// TIA Portal project "2026_09_21_Ciclo_L" (V15)

(* hardware
DEVICE "S7-1200 station_1"  S7-1200 Station
   slot 0: "Telaio di montaggio_0"  S7-1200 Rack  Rack  V1.0
   slot 1: "PLC_1"  CPU 1215C DC/DC/DC  6ES7 215-1AG40-0XB0  V4.2
*)

// ===== PLC "PLC_1"  CPU 1215C DC/DC/DC =====

VAR_GLOBAL   // PLC tag table "Tabella delle variabili standard"
   "IC" AT %I0.0 : Bool;   // Pulsante di inizio ciclo
   "FC" AT %I0.1 : Bool;   // Pulsante di fine ciclo
   "a0" AT %I0.2 : Bool;   // Fine corsa cilindro A chiuso
   "a1" AT %I0.3 : Bool;   // Fine corsa cilindro A aperto
   "b0" AT %I0.4 : Bool;   // Fine corsa cilindro B chiuso
   "b1" AT %I0.5 : Bool;   // Fine corsa cilindro B aperto
   "A+" AT %Q0.0 : Bool;   // Fase positiva cilindro A
   "A-" AT %Q0.1 : Bool;   // Fase negativa cilindro A
   "B+" AT %Q0.2 : Bool;   // Fase positiva cilindro B
   "B-" AT %Q0.3 : Bool;   // Fase negativa cilindro B
   "HL0" AT %Q0.4 : Bool;   // Lampada di segnalazione impianto spento
   "HL1" AT %Q0.5 : Bool;   // Lampada di segnalazione impianto acceso
   "P0" AT %M10.0 : Bool;   // Fase 0
   "P1" AT %M10.1 : Bool;   // Fase 1
   "P2" AT %M10.2 : Bool;   // Fase 2
   "P3" AT %M10.3 : Bool;   // Fase 3
   "P4" AT %M10.4 : Bool;   // Fase 4
   "IC_V" AT %M20.0 : Bool;   // Start virtuale
   "FC_V" AT %M20.1 : Bool;
   "a0_V" AT %M20.2 : Bool;
   "a1_V" AT %M20.3 : Bool;
   "b0_V" AT %M20.4 : Bool;
   "b1_V" AT %M20.5 : Bool;
END_VAR

FUNCTION "Controllo" : Void   // FC1, LAD
{ S7_Optimized_Access := 'TRUE' }
VERSION : 0.1
   VAR_TEMP   // added for the SCL form of the ladder/FBD networks
      _w1 : Bool;
   END_VAR
BEGIN

REGION Network 1: Fase 0
   // Alla pressione del pulsante di Start, si avvia il ciclo di lavoro (stato 1)
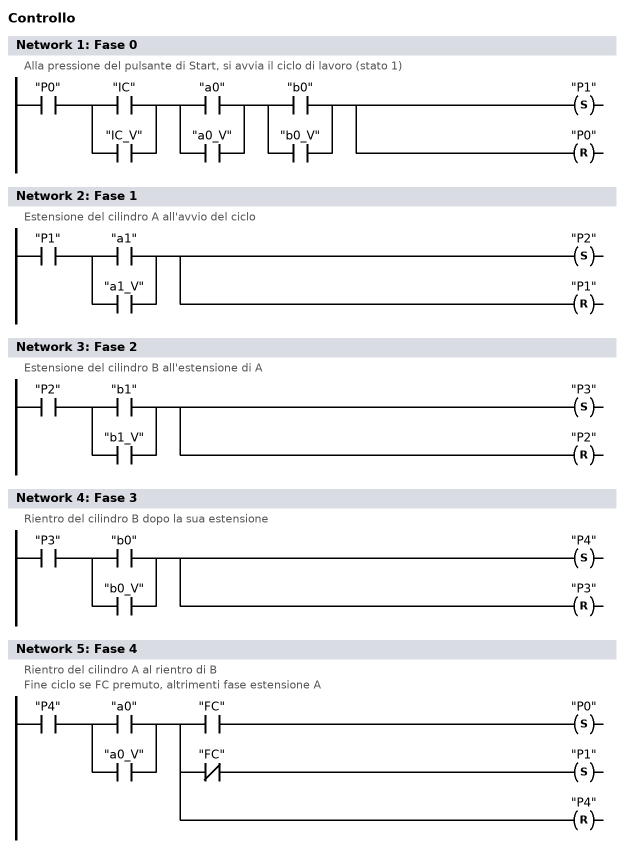
   RUNG wire#powerrail
      Contact( "P0" )
      wire#w1
      Contact( "IC" )
      wire#w2
      Contact( "a0" )
      wire#w3
      Contact( "b0" )
      wire#w4
      S_Coil( "P1" )
   END_RUNG
   RUNG wire#w1
      Contact( "IC_V" )
   END_RUNG wire#w2
   RUNG wire#w2
      Contact( "a0_V" )
   END_RUNG wire#w3
   RUNG wire#w3
      Contact( "b0_V" )
   END_RUNG wire#w4
   RUNG wire#w4
      R_Coil( "P0" )
   END_RUNG
   // the same network as SCL:
   IF "P0" AND ("IC" OR "IC_V") AND ("a0" OR "a0_V") AND ("b0" OR "b0_V") THEN
       "P1" := TRUE;
       "P0" := FALSE;
   END_IF;
END_REGION

REGION Network 2: Fase 1
   // Estensione del cilindro A all'avvio del ciclo
   RUNG wire#powerrail
      Contact( "P1" )
      wire#w1
      Contact( "a1" )
      wire#w2
      S_Coil( "P2" )
   END_RUNG
   RUNG wire#w1
      Contact( "a1_V" )
   END_RUNG wire#w2
   RUNG wire#w2
      R_Coil( "P1" )
   END_RUNG
   // the same network as SCL:
   IF "P1" AND ("a1" OR "a1_V") THEN
       "P2" := TRUE;
       "P1" := FALSE;
   END_IF;
END_REGION

REGION Network 3: Fase 2
   // Estensione del cilindro B all'estensione di A
   RUNG wire#powerrail
      Contact( "P2" )
      wire#w1
      Contact( "b1" )
      wire#w2
      S_Coil( "P3" )
   END_RUNG
   RUNG wire#w1
      Contact( "b1_V" )
   END_RUNG wire#w2
   RUNG wire#w2
      R_Coil( "P2" )
   END_RUNG
   // the same network as SCL:
   IF "P2" AND ("b1" OR "b1_V") THEN
       "P3" := TRUE;
       "P2" := FALSE;
   END_IF;
END_REGION

REGION Network 4: Fase 3
   // Rientro del cilindro B dopo la sua estensione
   RUNG wire#powerrail
      Contact( "P3" )
      wire#w1
      Contact( "b0" )
      wire#w2
      S_Coil( "P4" )
   END_RUNG
   RUNG wire#w1
      Contact( "b0_V" )
   END_RUNG wire#w2
   RUNG wire#w2
      R_Coil( "P3" )
   END_RUNG
   // the same network as SCL:
   IF "P3" AND ("b0" OR "b0_V") THEN
       "P4" := TRUE;
       "P3" := FALSE;
   END_IF;
END_REGION

REGION Network 5: Fase 4
   // Rientro del cilindro A al rientro di B
   // Fine ciclo se FC premuto, altrimenti fase estensione A
   RUNG wire#powerrail
      Contact( "P4" )
      wire#w1
      Contact( "a0" )
      wire#w2
      Contact( "FC" )
      S_Coil( "P0" )
   END_RUNG
   RUNG wire#w1
      Contact( "a0_V" )
   END_RUNG wire#w2
   RUNG wire#w2
      I_Contact( "FC" )
      S_Coil( "P1" )
   END_RUNG
   RUNG wire#w2
      R_Coil( "P4" )
   END_RUNG
   // the same network as SCL:
   #_w1 := "P4" AND ("a0" OR "a0_V");
   IF #_w1 AND "FC" THEN "P0" := TRUE; END_IF;
   IF #_w1 AND NOT "FC" THEN "P1" := TRUE; END_IF;
   IF #_w1 THEN "P4" := FALSE; END_IF;
END_REGION
END_FUNCTION

FUNCTION "Comando" : Void   // FC2, LAD
{ S7_Optimized_Access := 'TRUE' }
VERSION : 0.1
BEGIN

REGION Network 1: Lampada di segnalazione impianto spento
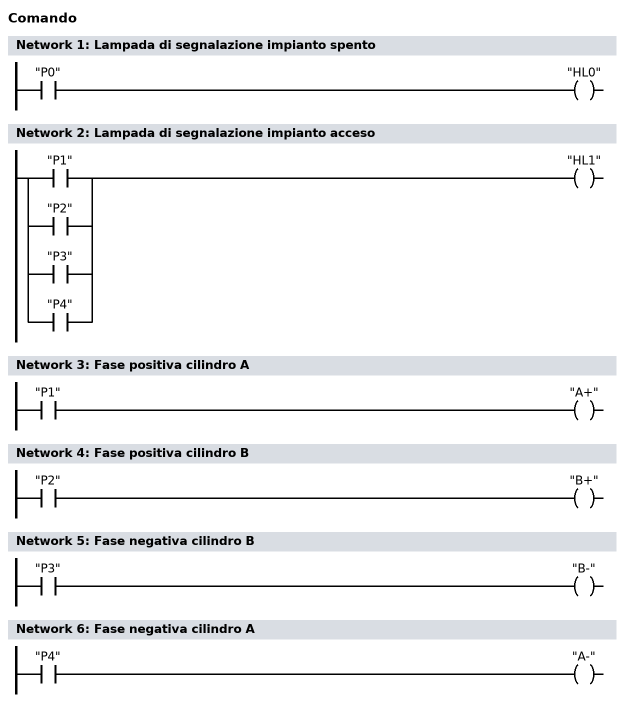
   RUNG wire#powerrail
      Contact( "P0" )
      Coil( "HL0" )
   END_RUNG
   // the same network as SCL:
   "HL0" := "P0";
END_REGION

REGION Network 2: Lampada di segnalazione impianto acceso
   RUNG wire#powerrail
      Contact( "P1" )
      wire#w1
      Coil( "HL1" )
   END_RUNG
   RUNG wire#powerrail
      Contact( "P2" )
   END_RUNG wire#w1
   RUNG wire#powerrail
      Contact( "P3" )
   END_RUNG wire#w1
   RUNG wire#powerrail
      Contact( "P4" )
   END_RUNG wire#w1
   // the same network as SCL:
   "HL1" := "P1" OR "P2" OR "P3" OR "P4";
END_REGION

REGION Network 3: Fase positiva cilindro A
   RUNG wire#powerrail
      Contact( "P1" )
      Coil( "A+" )
   END_RUNG
   // the same network as SCL:
   "A+" := "P1";
END_REGION

REGION Network 4: Fase positiva cilindro B
   RUNG wire#powerrail
      Contact( "P2" )
      Coil( "B+" )
   END_RUNG
   // the same network as SCL:
   "B+" := "P2";
END_REGION

REGION Network 5: Fase negativa cilindro B
   RUNG wire#powerrail
      Contact( "P3" )
      Coil( "B-" )
   END_RUNG
   // the same network as SCL:
   "B-" := "P3";
END_REGION

REGION Network 6: Fase negativa cilindro A
   RUNG wire#powerrail
      Contact( "P4" )
      Coil( "A-" )
   END_RUNG
   // the same network as SCL:
   "A-" := "P4";
END_REGION
END_FUNCTION

ORGANIZATION_BLOCK "Main"   // OB1, LAD, ProgramCycle
TITLE = "Main Program Sweep (Cycle)"
{ S7_Optimized_Access := 'TRUE' }
VERSION : 0.1
   VAR_INPUT
      Initial_Call : Bool;   // Initial call of this OB
      Remanence : Bool;   // =True, if remanent data are available
   END_VAR
BEGIN

REGION Network 1: FC Controllo
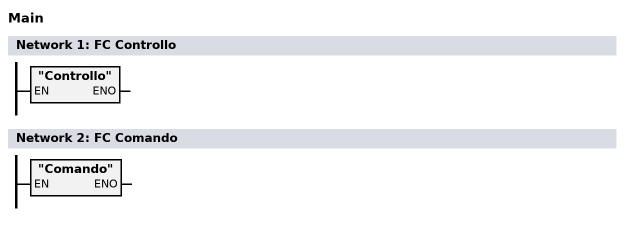
   RUNG wire#powerrail
      "Controllo"()
   END_RUNG
   // the same network as SCL:
   "Controllo"();
END_REGION

REGION Network 2: FC Comando
   RUNG wire#powerrail
      "Comando"()
   END_RUNG
   // the same network as SCL:
   "Comando"();
END_REGION
END_ORGANIZATION_BLOCK

ORGANIZATION_BLOCK "Startup"   // OB100, LAD, Startup
TITLE = "Complete Restart"
{ S7_Optimized_Access := 'TRUE' }
VERSION : 0.1
   VAR_INPUT
      LostRetentive : Bool;   // True if retentive data are lost
      LostRTC : Bool;   // True if date and time are lost
   END_VAR
BEGIN

REGION Network 1: Reset fasi
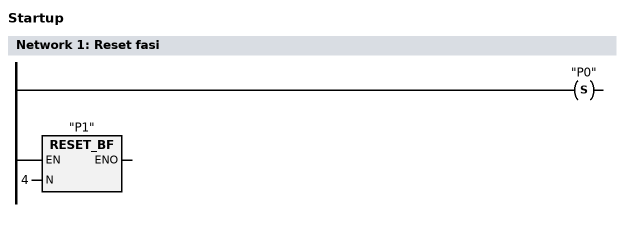
   // no SCL statement known for RBitfield: written as a call
   "P0" := TRUE;
   RESET_BF(operand := "P1", n := 4);
END_REGION
END_ORGANIZATION_BLOCK